// TIA Portal V20 export
// export: Created 2026-10-12T04:58:19.9885886Z, ExportSetting WithDefaults, DisplayName Totally Integrated Automation Portal, DisplayVersion V20, DisplayName TIA Portal Openness, DisplayVersion V20, DisplayName TIA Portal Teamcenter Gateway, DisplayVersion V20, DisplayName TIA Portal Version Control Interface, DisplayVersion V20, DisplayName SINAMICS Startdrive Advanced, DisplayVersion V20 SP1 Update 2, DisplayName SINAMICS Startdrive G110M, G120, G120C, G120D, G120P, G115D, DisplayVersion V20 SP1 Update 2, DisplayName SINAMICS Startdrive G130, G150, S120, S150, SINAMICS MV, G220, S200, S210, DisplayVersion V20 SP1 Update 2, DisplayName STEP 7 Professional, DisplayVersion V20, DisplayName STEP 7 Safety, DisplayVersion V20, DisplayName WinCC Basic/Comfort/Advanced, DisplayVersion V20, DisplayName WinCC Professional, DisplayVersion V20, DisplayName WinCC Unified, DisplayVersion V20
FUNCTION "FRK_AccessUsersShape" : Bool   // FC52, SCL
{ S7_Optimized_Access := 'TRUE' }
VERSION : 0.1
// stored: AutoNumber true, IsIECCheckEnabled false, SetENOAutomatically false, UDAEnableTagReadback false
   VAR_TEMP
      Slot : Int;
      Other : Int;
   END_VAR
BEGIN

   #FRK_AccessUsersShape := FALSE;
   IF "FRK_LocalUsers".Count < 0 OR "FRK_LocalUsers".Count > 16 THEN
       RETURN;
   END_IF;
   FOR #Slot := 1 TO DINT_TO_INT("FRK_LocalUsers".Count) DO
       IF "FRK_LocalUsers".Rows[#Slot].User = '' OR "FRK_LocalUsers".Rows[#Slot].Level < 1 OR "FRK_LocalUsers".Rows[#Slot].Level > 4 THEN
           RETURN;
       END_IF;
       FOR #Other := 1 TO #Slot - 1 DO
           IF "FRK_LocalUsers".Rows[#Slot].User = "FRK_LocalUsers".Rows[#Other].User THEN
               RETURN;
           END_IF;
       END_FOR;
   END_FOR;
   #FRK_AccessUsersShape := TRUE;
END_FUNCTION
